Fanuc KAREL source: KO00092.KL

PROGRAM KO00092
%NOLOCKGROUP
%ENVIRONMENT MIR
VAR
  P1: JOINTPOS
  P2: XYZWPREXT
  F: BOOLEAN
  OUT: JOINTPOS
BEGIN
  F = TRUE
  OUT = MIRROR(P1, P2, F)
END KO00092
